(* IEC 61131-3 sources: plcassist-cli/packages/volt-lsp-iec/test-corpus/CodesysTestProject/Device/Plc Logic/Application/Library Manager/CmpIoMgr Implementation, 47 files *)

(* ---- IOMGRCONFIGGETCONNECTOR.fun ---- *)
FUNCTION IOMGRCONFIGGETCONNECTOR : POINTER TO IoConfigConnector
VAR_INPUT
	PCONNECTORLIST : POINTER TO IoConfigConnector;
	PNCOUNT : POINTER TO DINT;
	DWMODULETYPE : DWORD;
	DWINSTANCE : DWORD;
END_VAR
END_FUNCTION

(* ---- IOMGRCONFIGGETCONNECTORBYDRIVER.fun ---- *)
FUNCTION IOMGRCONFIGGETCONNECTORBYDRIVER : POINTER TO IoConfigConnector
VAR_INPUT
	PIBASE : IBase;
	BIECDRIVER : DINT;
	NINDEX : DINT;
	PRESULT : POINTER TO RTS_IEC_RESULT;
END_VAR
END_FUNCTION

(* ---- IOMGRCONFIGGETCONNECTORLIST.fun ---- *)
FUNCTION IOMGRCONFIGGETCONNECTORLIST : RTS_IEC_RESULT
VAR_INPUT
	PPCONNECTORLIST : POINTER TO POINTER TO IoConfigConnector;
	PNCOUNT : POINTER TO DINT;
END_VAR
END_FUNCTION

(* ---- IOMGRCONFIGGETDRIVER.fun ---- *)
FUNCTION IOMGRCONFIGGETDRIVER : IBase
VAR_INPUT
	PCONNECTOR : POINTER TO IoConfigConnector;
	PBIECDRIVER : POINTER TO DINT;
	PRESULT : POINTER TO RTS_IEC_RESULT;
END_VAR
END_FUNCTION

(* ---- IOMGRCONFIGGETFIRSTCHILD.fun ---- *)
FUNCTION IOMGRCONFIGGETFIRSTCHILD : POINTER TO IoConfigConnector
VAR_INPUT
	PCONNECTORLIST : POINTER TO IoConfigConnector;
	PNCOUNT : POINTER TO DINT;
	PFATHER : POINTER TO IoConfigConnector;
END_VAR
END_FUNCTION

(* ---- IOMGRCONFIGGETFIRSTCONNECTOR.fun ---- *)
FUNCTION IOMGRCONFIGGETFIRSTCONNECTOR : POINTER TO IoConfigConnector
VAR_INPUT
	PCONNECTORLIST : POINTER TO IoConfigConnector;
	PNCOUNT : POINTER TO DINT;
	WTYPE : WORD;
END_VAR
END_FUNCTION

(* ---- IOMGRCONFIGGETNEXTCHILD.fun ---- *)
FUNCTION IOMGRCONFIGGETNEXTCHILD : POINTER TO IoConfigConnector
VAR_INPUT
	PCONNECTORLIST : POINTER TO IoConfigConnector;
	PNCOUNT : POINTER TO DINT;
	PFATHER : POINTER TO IoConfigConnector;
END_VAR
END_FUNCTION

(* ---- IOMGRCONFIGGETNEXTCONNECTOR.fun ---- *)
FUNCTION IOMGRCONFIGGETNEXTCONNECTOR : POINTER TO IoConfigConnector
VAR_INPUT
	PCONNECTORLIST : POINTER TO IoConfigConnector;
	PNCOUNT : POINTER TO DINT;
	WTYPE : WORD;
END_VAR
END_FUNCTION

(* ---- IOMGRCONFIGGETPARAMETER.fun ---- *)
FUNCTION IOMGRCONFIGGETPARAMETER : POINTER TO IoConfigParameter
VAR_INPUT
	PCONNECTOR : POINTER TO IoConfigConnector;
	DWPARAMETERID : DWORD;
END_VAR
END_FUNCTION

(* ---- IOMGRCONFIGGETPARAMETERVALUEBYTE.fun ---- *)
FUNCTION IOMGRCONFIGGETPARAMETERVALUEBYTE : BYTE
VAR_INPUT
	PPARAMETER : POINTER TO IoConfigParameter;
	PRESULT : POINTER TO UDINT;
END_VAR
END_FUNCTION

(* ---- IOMGRCONFIGGETPARAMETERVALUEDWORD.fun ---- *)
FUNCTION IOMGRCONFIGGETPARAMETERVALUEDWORD : DWORD
VAR_INPUT
	PPARAMETER : POINTER TO IoConfigParameter;
	PRESULT : POINTER TO UDINT;
END_VAR
END_FUNCTION

(* ---- IOMGRCONFIGGETPARAMETERVALUEPOINTER.fun ---- *)
FUNCTION IOMGRCONFIGGETPARAMETERVALUEPOINTER : POINTER TO BYTE
VAR_INPUT
	PPARAMETER : POINTER TO IoConfigParameter;
	PRESULT : POINTER TO UDINT;
END_VAR
END_FUNCTION

(* ---- IOMGRCONFIGGETPARAMETERVALUEWORD.fun ---- *)
FUNCTION IOMGRCONFIGGETPARAMETERVALUEWORD : WORD
VAR_INPUT
	PPARAMETER : POINTER TO IoConfigParameter;
	PRESULT : POINTER TO UDINT;
END_VAR
END_FUNCTION

(* ---- IOMGRCONFIGRESETDIAGNOSIS.fun ---- *)
FUNCTION IOMGRCONFIGRESETDIAGNOSIS : UDINT
VAR_INPUT
	PCONNECTOR : POINTER TO IoConfigConnector;
	DWFLAGS : DWORD;
END_VAR
END_FUNCTION

(* ---- IOMGRCONFIGSETDIAGNOSIS.fun ---- *)
FUNCTION IOMGRCONFIGSETDIAGNOSIS : UDINT
VAR_INPUT
	PCONNECTOR : POINTER TO IoConfigConnector;
	DWFLAGS : DWORD;
END_VAR
END_FUNCTION

(* ---- IOMGRCOPYINPUTBE.fun ---- *)
FUNCTION IOMGRCOPYINPUTBE : RTS_IEC_RESULT
VAR_INPUT
	PCHANNEL : POINTER TO IoConfigChannelMap;
	PADDRESS : POINTER TO BYTE;
END_VAR
END_FUNCTION

(* ---- IOMGRCOPYINPUTLE.fun ---- *)
FUNCTION IOMGRCOPYINPUTLE : RTS_IEC_RESULT
VAR_INPUT
	PCHANNEL : POINTER TO IoConfigChannelMap;
	PADDRESS : POINTER TO BYTE;
END_VAR
END_FUNCTION

(* ---- IOMGRCOPYOUTPUTBE.fun ---- *)
FUNCTION IOMGRCOPYOUTPUTBE : RTS_IEC_RESULT
VAR_INPUT
	PCHANNEL : POINTER TO IoConfigChannelMap;
	PADDRESS : POINTER TO BYTE;
END_VAR
END_FUNCTION

(* ---- IOMGRCOPYOUTPUTLE.fun ---- *)
FUNCTION IOMGRCOPYOUTPUTLE : RTS_IEC_RESULT
VAR_INPUT
	PCHANNEL : POINTER TO IoConfigChannelMap;
	PADDRESS : POINTER TO BYTE;
END_VAR
END_FUNCTION

(* ---- IOMGRGETBUSCYCLETYPE.fun ---- *)
FUNCTION IOMGRGETBUSCYCLETYPE : UDINT
VAR_INPUT
	PCONNECTOR : POINTER TO IoConfigConnector;
	PRESULT : POINTER TO RTS_IEC_RESULT;
END_VAR
END_FUNCTION

(* ---- IOMGRGETCONFIGAPPLICATION.fun ---- *)
FUNCTION IOMGRGETCONFIGAPPLICATION : RTS_IEC_RESULT
VAR_INPUT
	PSZCONFIGAPPLICATION : REFERENCE TO STRING;
	PNMAXLEN : POINTER TO DINT;
END_VAR
END_FUNCTION

(* ---- IOMGRGETDRIVERPROPERTIES.fun ---- *)
FUNCTION IOMGRGETDRIVERPROPERTIES : RTS_IEC_RESULT
VAR_INPUT
	HIODRV : RTS_IEC_HANDLE;
	PPPROPERTIES : POINTER TO POINTER TO DWORD;
END_VAR
END_FUNCTION

(* ---- IOMGRGETFIRSTDRIVERINSTANCE.fun ---- *)
FUNCTION IOMGRGETFIRSTDRIVERINSTANCE : IBase
VAR_INPUT
	PBIECDRIVER : POINTER TO DINT;
	PRESULT : POINTER TO RTS_IEC_RESULT;
END_VAR
END_FUNCTION

(* ---- IOMGRGETMODULEDIAGNOSIS.fun ---- *)
FUNCTION IOMGRGETMODULEDIAGNOSIS : UDINT
VAR_INPUT
	PCONNECTOR : POINTER TO IoConfigConnector;
END_VAR
END_FUNCTION

(* ---- IOMGRGETNEXTDRIVERINSTANCE.fun ---- *)
FUNCTION IOMGRGETNEXTDRIVERINSTANCE : IBase
VAR_INPUT
	PIBASEPREV : IBase;
	PBIECDRIVER : POINTER TO DINT;
	PRESULT : POINTER TO RTS_IEC_RESULT;
END_VAR
END_FUNCTION

(* ---- IOMGRIDENTIFY.fun ---- *)
FUNCTION IOMGRIDENTIFY : UDINT
VAR_INPUT
	PCONNECTOR : POINTER TO IoConfigConnector;
END_VAR
END_FUNCTION

(* ---- IOMGRLOCKENTER.fun ---- *)
FUNCTION IOMGRLOCKENTER : RTS_IEC_RESULT
VAR_INPUT
	HIODRV : RTS_IEC_HANDLE;
	DWLOCKSCOPE : DWORD;
END_VAR
END_FUNCTION

(* ---- IOMGRLOCKLEAVE.fun ---- *)
FUNCTION IOMGRLOCKLEAVE : RTS_IEC_RESULT
VAR_INPUT
	HIODRV : RTS_IEC_HANDLE;
	DWLOCKSCOPE : DWORD;
END_VAR
END_FUNCTION

(* ---- IOMGRREADINPUTS.fun ---- *)
FUNCTION IOMGRREADINPUTS : UDINT
VAR_INPUT
	PTASKMAP : POINTER TO IoConfigTaskMap;
END_VAR
END_FUNCTION

(* ---- IOMGRREADPARAMETER.fun ---- *)
FUNCTION IOMGRREADPARAMETER : UDINT
VAR_INPUT
	DWMODULETYPE : DWORD;
	DWINSTANCE : DWORD;
	DWPARAMETERID : DWORD;
	PDATA : POINTER TO BYTE;
	DWBITSIZE : DWORD;
	DWBITOFFSET : DWORD;
END_VAR
END_FUNCTION

(* ---- IOMGRRECONFIGURE.fun ---- *)
FUNCTION IOMGRRECONFIGURE : RTS_IEC_RESULT
VAR_INPUT
	PCONNECTOR : POINTER TO IoConfigConnector;
	PUDISTATE : POINTER TO UDINT;
END_VAR
END_FUNCTION

(* ---- IOMGRREGISTERCONFIGAPPLICATION.fun ---- *)
FUNCTION IOMGRREGISTERCONFIGAPPLICATION : RTS_IEC_RESULT
VAR_INPUT
	PSZCONFIGAPPLICATION : REFERENCE TO STRING;
END_VAR
END_FUNCTION

(* ---- IOMGRREGISTERINSTANCE2.fun ---- *)
FUNCTION IOMGRREGISTERINSTANCE2 : RTS_IEC_HANDLE
VAR_INPUT
	DWCLASSID : DWORD;
	PITF : IBase;
	PRESULT : POINTER TO RTS_IEC_RESULT;
END_VAR
END_FUNCTION

(* ---- IOMGRSCANMODULES.fun ---- *)
FUNCTION IOMGRSCANMODULES : UDINT
VAR_INPUT
	PCONNECTOR : POINTER TO IoConfigConnector;
	PPCONNECTORLIST : POINTER TO POINTER TO IoConfigConnector;
	PNCOUNT : POINTER TO DINT;
END_VAR
END_FUNCTION

(* ---- IOMGRSETDRIVERPROPERTIES.fun ---- *)
FUNCTION IOMGRSETDRIVERPROPERTIES : RTS_IEC_RESULT
VAR_INPUT
	HIODRV : RTS_IEC_HANDLE;
	ULPROPERTIES : DWORD;
END_VAR
END_FUNCTION

(* ---- IOMGRSETDRIVERPROPERTY.fun ---- *)
FUNCTION IOMGRSETDRIVERPROPERTY : RTS_IEC_RESULT
VAR_INPUT
	HIODRV : RTS_IEC_HANDLE;
	ULPROPERTY : DWORD;
	BVALUE : DINT;
END_VAR
END_FUNCTION

(* ---- IOMGRSTARTBUSCYCLE.fun ---- *)
FUNCTION IOMGRSTARTBUSCYCLE : UDINT
VAR_INPUT
	PCONNECTOR : POINTER TO IoConfigConnector;
END_VAR
END_FUNCTION

(* ---- IOMGRSTARTBUSCYCLE2.fun ---- *)
FUNCTION IOMGRSTARTBUSCYCLE2 : UDINT
VAR_INPUT
	PCONNECTOR : POINTER TO IoConfigConnector;
	DWTYPE : UDINT;
END_VAR
END_FUNCTION

(* ---- IOMGRUNREGISTERCONFIGAPPLICATION.fun ---- *)
FUNCTION IOMGRUNREGISTERCONFIGAPPLICATION : RTS_IEC_RESULT
VAR_INPUT
	PSZCONFIGAPPLICATION : REFERENCE TO STRING;
END_VAR
END_FUNCTION

(* ---- IOMGRUNREGISTERINSTANCE.fun ---- *)
FUNCTION IOMGRUNREGISTERINSTANCE : RTS_IEC_RESULT
VAR_INPUT
	HINTERFACE : RTS_IEC_HANDLE;
END_VAR
END_FUNCTION

(* ---- IOMGRUPDATECONFIGURATION.fun ---- *)
FUNCTION IOMGRUPDATECONFIGURATION : UDINT
VAR_INPUT
	PCONNECTORLIST : POINTER TO IoConfigConnector;
	NCOUNT : DINT;
END_VAR
END_FUNCTION

(* ---- IOMGRUPDATECONFIGURATION2.fun ---- *)
FUNCTION IOMGRUPDATECONFIGURATION2 : UDINT
VAR_INPUT
	PCONNECTORLIST : POINTER TO IoConfigConnector;
	NCOUNT : DINT;
	PSZCONFIGAPPLICATION : REFERENCE TO STRING;
END_VAR
END_FUNCTION

(* ---- IOMGRUPDATEMAPPING.fun ---- *)
FUNCTION IOMGRUPDATEMAPPING : UDINT
VAR_INPUT
	PTASKMAPLIST : POINTER TO IoConfigTaskMap;
	NCOUNT : DINT;
END_VAR
END_FUNCTION

(* ---- IOMGRUPDATEMAPPING2.fun ---- *)
FUNCTION IOMGRUPDATEMAPPING2 : UDINT
VAR_INPUT
	PTASKMAPLIST : POINTER TO IoConfigTaskMap;
	NCOUNT : DINT;
	PSZCONFIGAPPLICATION : REFERENCE TO STRING;
END_VAR
END_FUNCTION

(* ---- IOMGRWATCHDOGTRIGGER.fun ---- *)
FUNCTION IOMGRWATCHDOGTRIGGER : UDINT
VAR_INPUT
	PCONNECTOR : POINTER TO IoConfigConnector;
END_VAR
END_FUNCTION

(* ---- IOMGRWRITEOUTPUTS.fun ---- *)
FUNCTION IOMGRWRITEOUTPUTS : UDINT
VAR_INPUT
	PTASKMAP : POINTER TO IoConfigTaskMap;
END_VAR
END_FUNCTION

(* ---- IOMGRWRITEPARAMETER.fun ---- *)
FUNCTION IOMGRWRITEPARAMETER : UDINT
VAR_INPUT
	DWMODULETYPE : DWORD;
	DWINSTANCE : DWORD;
	DWPARAMETERID : DWORD;
	PDATA : POINTER TO BYTE;
	DWBITSIZE : DWORD;
	DWBITOFFSET : DWORD;
END_VAR
END_FUNCTION
